TYPE ST_PersistentWriteRequest :
STRUCT
	ModuleId : UDINT;
	ServiceId : UDINT;
END_STRUCT
END_TYPE

(* stored: Version 1.1.0.1, ProductVersion 3.1.4026.18
   DUT ST_PersistentWriteRequest: Id {7feac50f-a753-45d8-8aa5-0904f173c5f1} *)
